(* IEC 61131-3 sources: kns-pump-station/tests/POUs/Station/FB_F_StationCfgCheck_Test, 13 files *)

(* ---- AlarmBit.method.decl.st ---- *)
// 04 §18.3: приоритет тревоги станции вне перечисления — STN_CFG_ALARM
METHOD PRIVATE AlarmBit
VAR
    stCfg : ST_StationCfg;              // уставки по умолчанию (04 §18.2)
    stPid : PL.ST_PidCfg;               // LIC101: пределы задания 1,2…2,2 м
    wErr  : WORD;                       // результат проверки
    pRaw : POINTER TO INT;           // значение вне перечисления
END_VAR

(* ---- DefaultsPass.method.decl.st ---- *)
// 04 §18.2: уставки по умолчанию с отметками L 0,8 м и H 3,5 м проходят проверку
METHOD PRIVATE DefaultsPass
VAR
    stCfg : ST_StationCfg;              // уставки по умолчанию (04 §18.2)
    stPid : PL.ST_PidCfg;               // LIC101: пределы задания 1,2…2,2 м
    wErr  : WORD;                       // результат проверки
END_VAR

(* ---- DutyBit.method.decl.st ---- *)
// 04 §18.2 № 13: uiDutyMax вне 1…3 — STN_CFG_DUTY
METHOD PRIVATE DutyBit
VAR
    stCfg : ST_StationCfg;              // уставки по умолчанию (04 §18.2)
    stPid : PL.ST_PidCfg;               // LIC101: пределы задания 1,2…2,2 м
    wErr  : WORD;                       // результат проверки
END_VAR

(* ---- FloatCheckBit.method.decl.st ---- *)
// 04 §18.2 № 22–26: отметки и выдержка согласования поплавков вне диапазонов — STN_CFG_FLOAT_CHECK
METHOD PRIVATE FloatCheckBit
VAR
    stCfg : ST_StationCfg;              // уставки по умолчанию (04 §18.2)
    stPid : PL.ST_PidCfg;               // LIC101: пределы задания 1,2…2,2 м
    wErr  : WORD;                       // результат проверки
END_VAR

(* ---- LevelOrderBit.method.decl.st ---- *)
// 04 §1, PMI-08 шаг 3: нарушен порядок отметок (останов подпорного выше пуска ведущего; H ниже пуска подпорного) —
// STN_CFG_LEVEL_ORDER
METHOD PRIVATE LevelOrderBit
VAR
    stCfg : ST_StationCfg;              // уставки по умолчанию (04 §18.2)
    stPid : PL.ST_PidCfg;               // LIC101: пределы задания 1,2…2,2 м
    wErr  : WORD;                       // результат проверки
END_VAR

(* ---- LevelRangeBit.method.decl.st ---- *)
// 04 §18.2 № 2–5: уровень вне диапазона или зазор пуска меньше 0,3 м — STN_CFG_LEVEL_RANGE; ровно 0,3 м —
// допустимо
METHOD PRIVATE LevelRangeBit
VAR
    stCfg : ST_StationCfg;              // уставки по умолчанию (04 §18.2)
    stPid : PL.ST_PidCfg;               // LIC101: пределы задания 1,2…2,2 м
    wErr  : WORD;                       // результат проверки
END_VAR

(* ---- NanRejected.method.decl.st ---- *)
// 04 §18.3: неконечные уставки (NaN) не проходят проверки своих групп
METHOD PRIVATE NanRejected
VAR
    stCfg : ST_StationCfg;              // уставки по умолчанию (04 §18.2)
    stPid : PL.ST_PidCfg;               // LIC101: пределы задания 1,2…2,2 м
    wErr  : WORD;                       // результат проверки
    uBits : PL.U_RealBits;            // сборка NaN по битам
END_VAR

(* ---- PidStagingBit.method.decl.st ---- *)
// 04 §18.2 № 9–12, §18.3: rAssistOff_pct <= rAssistOn_pct - 10 (ровно — допустимо), выдержки в диапазоне — иначе
// STN_CFG_PID_STAGING
METHOD PRIVATE PidStagingBit
VAR
    stCfg : ST_StationCfg;              // уставки по умолчанию (04 §18.2)
    stPid : PL.ST_PidCfg;               // LIC101: пределы задания 1,2…2,2 м
    wErr  : WORD;                       // результат проверки
END_VAR

(* ---- RotationBit.method.decl.st ---- *)
// 04 §18.2 № 14–17: режим чередования вне перечисления, tMaxContRun между 0 и 10 мин — STN_CFG_ROTATION; 0 —
// выключено, допустимо
METHOD PRIVATE RotationBit
VAR
    stCfg : ST_StationCfg;              // уставки по умолчанию (04 §18.2)
    stPid : PL.ST_PidCfg;               // LIC101: пределы задания 1,2…2,2 м
    wErr  : WORD;                       // результат проверки
    pRaw : POINTER TO INT;           // значение вне перечисления
END_VAR

(* ---- SetpointBit.method.decl.st ---- *)
// 04 §18.2 № 8, PMI-08 шаг 2: задание уровня вне пределов задания LIC101 — STN_CFG_SETPOINT
METHOD PRIVATE SetpointBit
VAR
    stCfg : ST_StationCfg;              // уставки по умолчанию (04 §18.2)
    stPid : PL.ST_PidCfg;               // LIC101: пределы задания 1,2…2,2 м
    wErr  : WORD;                       // результат проверки
END_VAR

(* ---- SpeedBit.method.decl.st ---- *)
// 04 §18.2 № 7: частота ступенчатого режима вне 60…100 % — STN_CFG_SPEED
METHOD PRIVATE SpeedBit
VAR
    stCfg : ST_StationCfg;              // уставки по умолчанию (04 §18.2)
    stPid : PL.ST_PidCfg;               // LIC101: пределы задания 1,2…2,2 м
    wErr  : WORD;                       // результат проверки
END_VAR

(* ---- TimesBit.method.decl.st ---- *)
// 04 §18.2 № 6, 18–21, 27, 31: выдержки вне диапазонов — STN_CFG_TIMES
METHOD PRIVATE TimesBit
VAR
    stCfg : ST_StationCfg;              // уставки по умолчанию (04 §18.2)
    stPid : PL.ST_PidCfg;               // LIC101: пределы задания 1,2…2,2 м
    wErr  : WORD;                       // результат проверки
END_VAR

(* ---- UnderloadBit.method.decl.st ---- *)
// 04 §18.2 № 28–30: порог тока выше 30 А — STN_CFG_UNDERLOAD; 0 (выключено) — допустимо
METHOD PRIVATE UnderloadBit
VAR
    stCfg : ST_StationCfg;              // уставки по умолчанию (04 §18.2)
    stPid : PL.ST_PidCfg;               // LIC101: пределы задания 1,2…2,2 м
    wErr  : WORD;                       // результат проверки
END_VAR
